// TIA Portal V21 export
// export: Created 2026-11-10T07:35:02.9312982Z, ExportSetting WithDefaults, DisplayName Totally Integrated Automation Portal, DisplayVersion V21 Update 3, DisplayName STEP 7 Professional, DisplayVersion V21 Update 3, DisplayName STEP 7 Safety, DisplayVersion V21, DisplayName Tech WebApplication, DisplayVersion V21, DisplayName WinCC Basic/Comfort/Advanced, DisplayVersion V21 Update 3, DisplayName WinCC Unified, DisplayVersion V21 Update 3
FUNCTION_BLOCK "FB_Lad_ex025"   // FB64, LAD
{ S7_Optimized_Access := 'TRUE' }
VERSION : 0.1
// stored: AutoNumber true, IsIECCheckEnabled false, IsRetainMemResEnabled false, MemoryReserve 100, SetENOAutomatically false, UDAEnableTagReadback false
   VAR_INPUT
      v_n : Int;
      v_ret_val : Word;
   END_VAR
   VAR_IN_OUT
      v_in : Variant;
      v_out : Variant;
   END_VAR
BEGIN

REGION Network 1: ATH - Convert ASCII string to hexadecimal number
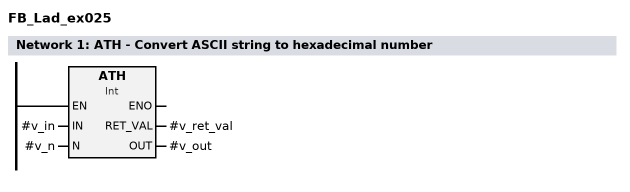
   RUNG wire#powerrail
      { S7_Templates := "[n_type := Int, in_out_type := Variant]" } ATH(IN := #v_in, N := #v_n, RET_VAL => #v_ret_val, OUT => #v_out)
   END_RUNG
   // the same network as SCL:
   #v_ret_val := ATH(IN := #v_in, N := #v_n, OUT => #v_out);
END_REGION
END_FUNCTION_BLOCK
